{attribute 'qualified_only'}
{attribute 'strict'}
TYPE E_EsolutionControl : (
	EmergencyShutdown := 11,
	SystemContactor := 12,	// 40013 Rack Contactor Control (맵 v1.4 이름): 1이면 랙 8개가 40001과 상관없이 한꺼번에 붙음
	ChargeContactor := 13,
	DischargeContactor := 14,
	ResetSystem := 30	// 40031 Reset System: 1이면 비상차단 해제 (명세 WR-BAT-01 v2.34)
) INT;
END_TYPE

(* stored: Version 1.1.0.1, ProductVersion 3.1.4024.15
   DUT E_EsolutionControl: Id {e57cb7c1-a0f5-46f0-877c-93d8f0d593ed} *)
